Fanuc KAREL source: ka00011.KL

-- PROVISIONAL review KL for V940-1; original PC SHA256 ecf77d44b28e2a19435701c084d7b6b6b708e77da65a25c7a4a69ed5ae85e53c
-- Incomplete behavior may be omitted. Consult companion uncertainty JSON. Do not deploy.
PROGRAM KA00011
%NOLOCKGROUP
VAR
  SRC : INTEGER
-- UNRESOLVED_DECL DST type=002018
BEGIN
  -- V9_ZERO_TABLE_METADATA_HINT layout=0001; no indexed target words; source/name/runtime held
  -- UNRESOLVED_PC offsets 5-16; opcodes 2E,23
  -- UNRESOLVED_PC offsets 21-36; opcodes 21,22,9D,33,B2
  -- UNRESOLVED_PC offsets 41-45; opcodes 7F
END KA00011
